// TIA Portal V14 SP1 export
// export: Created 2000-01-01T00:00:00.0000000Z, ExportSetting None
FUNCTION "FC_Rung" : Void   // FC42, LAD
{ S7_Optimized_Access := 'TRUE' }
   VAR_INPUT
      Local : Int;
   END_VAR
BEGIN

REGION Network 1
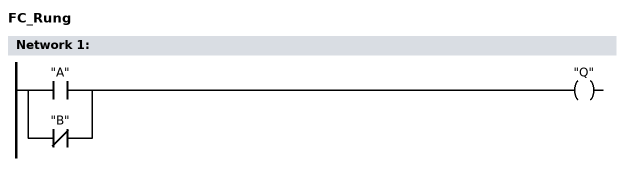
   RUNG wire#powerrail
      Contact( "A" )
      wire#w1
      Coil( "Q" )
   END_RUNG
   RUNG wire#powerrail
      I_Contact( "B" )
   END_RUNG wire#w1
   // the same network as SCL:
   "Q" := "A" OR NOT "B";
END_REGION
END_FUNCTION
